FUNCTION_BLOCK FB_STOEBERSI6SC6CIA402_REF
VAR_INPUT
	stTerminalState			AT %I*:ST_TerminalState;
	stStoeberToPlc			AT %I*:ST_STOEBERSI6SC6CIA402TOPLC;
	stPlcToStoeber			AT %Q*:ST_PLCTOSTOEBERSI6SC6CIA402;
END_VAR
VAR_OUTPUT

END_VAR
VAR_IN_OUT

END_VAR
VAR

END_VAR

;

END_FUNCTION_BLOCK

(* stored: Version 1.1.0.1, ProductVersion 3.1.4024.15
   POU FB_STOEBERSI6SC6CIA402_REF: Id {711d95d2-6373-4eae-8588-7dc9c1194d97}, SpecialFunc None *)
